FUNCTION_BLOCK FB_LeadLag (* Migrated from IEC 61131-3 ST *)
  (* Standard: 61499-2 *)
  (* Version 1.0, 2026-11-06, st2fb *)
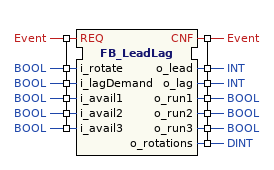
  EVENT_INPUT
    REQ WITH i_rotate, i_lagDemand, i_avail1, i_avail2, i_avail3;
  END_EVENT
  EVENT_OUTPUT
    CNF WITH o_lead, o_lag, o_run1, o_run2, o_run3, o_rotations;
  END_EVENT
  VAR_INPUT
    i_rotate : BOOL;
    i_lagDemand : BOOL;
    i_avail1 : BOOL;
    i_avail2 : BOOL;
    i_avail3 : BOOL;
  END_VAR
  VAR_OUTPUT
    o_lead : INT;
    o_lag : INT;
    o_run1 : BOOL;
    o_run2 : BOOL;
    o_run3 : BOOL;
    o_rotations : DINT;
  END_VAR
  VAR
    av1 : BOOL := FALSE;
    av2 : BOOL := FALSE;
    av3 : BOOL := FALSE;
    rot_Q : BOOL := FALSE;
    rot_M : BOOL := FALSE;
    tempIdx : INT := 0;
    tempCandidate : INT := 0;
    tempOffset : INT := 0;
    curAv : BOOL := FALSE;
    idxAv : BOOL := FALSE;
    done : BOOL := FALSE;
  END_VAR
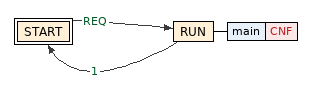
  EC_STATES
    START;
    RUN : main -> CNF;
  END_STATES
  EC_TRANSITIONS
    START TO RUN := REQ;
    RUN TO START := 1;
  END_TRANSITIONS
  ALGORITHM main IN ST:
av1 := i_avail1;
av2 := i_avail2;
av3 := i_avail3;

rot_Q := i_rotate AND NOT rot_M;
rot_M := i_rotate;

IF MAX(o_lead, 1) = 1 THEN
  curAv := av1;
ELSIF MAX(o_lead, 1) = 2 THEN
  curAv := av2;
ELSE
  curAv := av3;
END_IF;

IF rot_Q OR o_lead = 0 OR NOT curAv THEN
  tempCandidate := 0;
  done := FALSE;
  tempOffset := 1;
  WHILE tempOffset <= 3 AND NOT done DO
    tempIdx := (o_lead + tempOffset - 1) MOD 3 + 1;
    IF tempIdx = 1 THEN
      idxAv := av1;
    ELSIF tempIdx = 2 THEN
      idxAv := av2;
    ELSE
      idxAv := av3;
    END_IF;
    IF idxAv THEN
      tempCandidate := tempIdx;
      done := TRUE;
    END_IF;
    tempOffset := tempOffset + 1;
  END_WHILE;
  IF tempCandidate <> o_lead THEN
    o_lead := tempCandidate;
    o_rotations := o_rotations + 1;
  END_IF;
END_IF;

o_lag := 0;
IF i_lagDemand AND o_lead <> 0 THEN
  done := FALSE;
  tempOffset := 1;
  WHILE tempOffset <= 2 AND NOT done DO
    tempIdx := (o_lead + tempOffset - 1) MOD 3 + 1;
    IF tempIdx = 1 THEN
      idxAv := av1;
    ELSIF tempIdx = 2 THEN
      idxAv := av2;
    ELSE
      idxAv := av3;
    END_IF;
    IF idxAv THEN
      o_lag := tempIdx;
      done := TRUE;
    END_IF;
    tempOffset := tempOffset + 1;
  END_WHILE;
END_IF;

o_run1 := o_lead = 1 OR o_lag = 1;
o_run2 := o_lead = 2 OR o_lag = 2;
o_run3 := o_lead = 3 OR o_lag = 3;
  END_ALGORITHM
END_FUNCTION_BLOCK
